LAYER Default
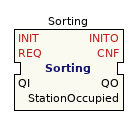
  FBS
    Sorting : Sorting;
  END_FBS
END_LAYER
